{attribute 'qualified_only'}
//{attribute 'strict'}
{attribute 'to_string'}
TYPE E_Pis_Name :
(
	e0_not_in_use := 0,
	// CIP Source
	V1001,
	V1002,
	V1003,
	V1004,
	V1005,

	MV1001,
	MV1002,
	MV1003,
	MV1004,
	
	//CIP Return
	V1101,
	V1102,
	V1103,
	V1104,
	V1105,
	V1112,
	V1114,
	V1117,
	V1120,
	
	//CIP Client
	V1106,
	V1023,V1024,V1025,V1026,V1027,V1028,V1029,V1030,

	//CIP Client Tanks
	V3001,V3003,V3005,V3006,V3007,V3041,V3039,
	V4001,V4003,V4005,V4006,V4007,V4041,V4039,	
	
	//CIP Tanks
	V1011,V1012,V1013,
	V1014,V1015,V1016,
	V1017,V1018,V1019,
	V1020,V1021,V1022,
	V1031,V1032,
	
	//Tank Target 1
	V3016,
	V3017,
	V3023,
	V3024,
	V3025,
	V3026,	
	
	//Tank Target 2
	V3015,	
	V3027,	
	V3028,	
	V3029,	
	V3030,	
	
	//Marinade Lines
	V3018,
	V3019,
	V3020,V3040,
	V3021,
	V3022,
	
	V3014,
	V3113,
	
	
	
	//Tank Target 3
	V4016,
	V4017,
	V4023,
	V4024,
	V4025,
	
	//Tank Target 4
	V4015,
	V4026,
	V4027,
	V4028,
	V4029,
	V4030,
	
	//Color Lines
	V4018,
	V4019,
	V4020,V4040,
	V4021,
	V4022,
	
	V2115,
	V2116,
	V2117,
	
	// Tanks Coolant
	V3031,V3032,
	V3033,V3034,
	V4031,V4032,
	V4042,V4043,
	
	//TriBlender Select
	V3035,V4037,V5001,
	V3038,V4038,V5002,
	
	//addition
	
	V4014,
	V4113,
	V2114,
	
	V3004,
	V3008,
	V3009,
	V3010,
	
	V4034,
	V4033,
	V4035,
	V4036,
	
	V4004,
	V4010,
	V4008,
	V4009,
	
	//Water
	V2011,V2111,V2211,V2112,
	
	
	V5012,
	
	V4026_2, //temp for marinade filling test 
	
	//Dummy valves for fbLineTarget_Marinade
	V_Dummy_01,
	V_Dummy_02,
	V_Dummy_03,
	V_Dummy_04,
	V_Dummy_05,
	V_Dummy_06,
	V_Dummy_07,
	V_Dummy_08,
	V_Dummy_09,
	V_Dummy_10,
	V_Dummy_11,
	V_Dummy_12,
	
	//Dummy for Line Source Marinada
	V_Dummy_LSM_01,
	V_Dummy_LSM_02,
	V_Dummy_LSM_03,
	V_Dummy_LSM_04,
	V_Dummy_LSM_05,
	V_Dummy_LSM_06,
	V_Dummy_LSM_07, //*
	//Dummy for TriBlender Source Marinada
	V_Dummy_TSM_01,
	V_Dummy_TSM_02,
	V_Dummy_TSM_03,
	//Dummy for Line Source Color
	V_Dummy_LSC_01,
	V_Dummy_LSC_02,
	V_Dummy_LSC_03,
	V_Dummy_LSC_04, //*
	
	//Dummy Drain Tap Water
	V_Dummy_DTW_01,
	
	
	//virtual list
	last
	



	
);
END_TYPE

(* stored: Version 1.1.0.1, ProductVersion 3.1.4024.15
   DUT E_Pis_Name: Id {c150e2d1-4733-4c0a-8dd7-5b1d3d1d7eff} *)
